Fanuc KAREL source: KT00219.KL

PROGRAM KT00219
%NOLOCKGROUP
VAR
  H1: ARRAY[2] OF SHORT
  I2: INTEGER
  OUT: BOOLEAN
BEGIN
  H1[1] = 2
    I2 = 3
  OUT = H1[1] AND I2
END KT00219
